(*
SPDX-FileCopyrightText: © 2026 Oleksandr Tiutyk <trofimich@gmail.com>
SPDX-License-Identifier: MIT
License: https://opensource.org/license/mit
*)

(*!
<summary>Exposes a scalar sort key for the collection natural-order fixture.</summary>
<description>
Borrowed interface used to reject unrelated IComparable implementations before reading a sort key.
</description>
*)

INTERFACE ICollectionSortValue EXTENDS TOF_Core.IComparable

(*!
<summary>Returns a copy of the fixture sort key without changing state.</summary>
*)
METHOD GetSortValue : DINT
END_METHOD

END_INTERFACE

(* stored: Version 1.1.0.1
   Itf ICollectionSortValue: Id {8beb5a96-aa8d-4024-9a3b-1936950af3d8}
   Method GetSortValue: Id {85a33168-1ff8-4a23-a9a0-cdbbdfe89c4f} *)
